SUBAPPLICATION Vorsteuerventil (* Subapplication Type *)
  (* Standard: 61499-2 *)
  (* Version 1.0, 2023-01-29, Franz *)
  IMPORT DataPanel::io::MI::DQ::DataPanel_MI_DO::Invalid;
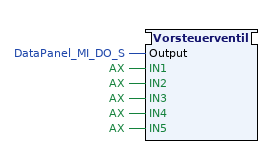
  VAR_INPUT
    Output : DataPanel::io::MI::DQ::DataPanel_MI_DO_S := Invalid;
  END_VAR
  SOCKETS
    IN1 : adapter::types::unidirectional::AX;
    IN2 : adapter::types::unidirectional::AX;
    IN3 : adapter::types::unidirectional::AX;
    IN4 : adapter::types::unidirectional::AX;
    IN5 : adapter::types::unidirectional::AX;
  END_SOCKETS
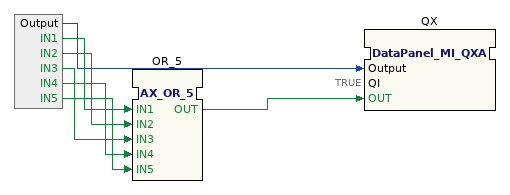
  FBS
    OR_5 : adapter::booleanOperators::AX_OR_5;
    QX : DataPanel::io::MI::DQ::DataPanel_MI_QXA(QI := TRUE);
  END_FBS
  DATA_CONNECTIONS
    Output TO QX.Output;
  END_CONNECTIONS
  ADAPTER_CONNECTIONS
    IN1 TO OR_5.IN1;
    IN2 TO OR_5.IN2;
    IN3 TO OR_5.IN3;
    IN4 TO OR_5.IN4;
    IN5 TO OR_5.IN5;
    OR_5.OUT TO QX.OUT;
  END_CONNECTIONS
END_SUBAPPLICATION
